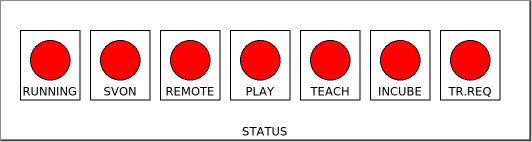
VISUALIZATION NX100_STATUS  // 532x142
    Rectangle (0,0 530x140), "STATUS"
    Rectangle (90,30 60x70), "SVON"
    Ellipse (100,40 40x40), colour toggle: MAIN.RSTATS.STATUS.ServoON
    Rectangle (160,30 60x70), "REMOTE"
    Ellipse (170,40 40x40), colour toggle: MAIN.RSTATS.STATUS.CommandRemote
    Rectangle (230,30 60x70), "PLAY"
    Ellipse (240,40 40x40), colour toggle: MAIN.RSTATS.STATUS.Play
    Rectangle (300,30 60x70), "TEACH"
    Ellipse (310,40 40x40), colour toggle: MAIN.RSTATS.STATUS.Teach
    Rectangle (370,30 60x70), "INCUBE"
    Ellipse (380,40 40x40), colour toggle: MAIN.InCube
    Rectangle (440,30 60x70), "TR.REQ"
    Ellipse (450,40 40x40), colour toggle: MAIN.TravelRequest
    Rectangle (20,30 60x70), "RUNNING"
    Ellipse (30,40 40x40), colour toggle: MAIN.RSTATS.STATUS.Running
END_VISUALIZATION

(* stored: Version 1.1.0.1, ProductVersion 3.1.4024.16
   Visu NX100_STATUS: Id {9694e602-947b-49cb-9fb2-df522eaf26a3} *)
